FUNCTION_BLOCK FB_LJ_S8000Capture
VAR_INPUT
	bExecute	:	BOOL	:=	FALSE;
END_VAR
VAR_OUTPUT
	bBusy		:	BOOL	:=	FALSE;
END_VAR
VAR
	nState		:	UDINT	:=	0;
END_VAR

CASE nState	OF

0:	
	IF bExecute	THEN
		IF NOT ExtPort.LJ_S8000_bTRG_ack THEN
			ExtPort.LJ_S8000_bTRG	:=	TRUE;
			bBusy	:=	TRUE;
			nState	:=	1;
		END_IF
	END_IF

1:
	IF ExtPort.LJ_S8000_bTRG_ack THEN
		ExtPort.LJ_S8000_bTRG	:=	FALSE;
	END_IF
	IF ExtPort.LJ_S8000_bBusy THEN
		nState	:=	2;
	END_IF
	
2:
	IF ExtPort.LJ_S8000_bReady THEN
		bBusy	:=	FALSE;
		nState	:=	0;
	END_IF
	
END_CASE

END_FUNCTION_BLOCK

(* stored: Version 1.1.0.1, ProductVersion 3.1.4024.15
   POU FB_LJ_S8000Capture: Id {969c9b00-c5ae-47a5-91f0-c2316712753f}, SpecialFunc None *)
